SUBAPPLICATION Button_IXA_OR_AX_BG (* Button (IXA) ODER AX-Eingang, Ergebnis als Hintergrundfarbe (Gruen/Weiss) und AX-Ausgang *)
  (* Standard: 61499-2; Description: Copyright (c) 2026 Meisterschulen am Ostbahnhof This program and the accompanying materials are made available under the terms of the Eclipse Public License 2.0 which is available at https://www.eclipse.org/legal/epl-2.0/ SPDX-License-Identifier: EPL-2.0 *)
  (* Version 1.0, 2026-10-31, Franz Höpfinger, Meisterschulen am Ostbahnhof, Aus Getreidehacke func/Manual/ManFuncTast0 in MyLib::sys verschoben und umbenannt, INIT/INITO/QI/QO ergaenzt. *)
  PACKAGE MyLib::sys;
  IMPORT isobus::UT::Q::const::IDs::ID_NULL;
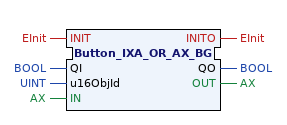
  EVENT_INPUT
    INIT : EInit; (* Initialization Request *)
  END_EVENT
  EVENT_OUTPUT
    INITO : EInit; (* Initialization Confirm *)
  END_EVENT
  VAR_INPUT
    QI : BOOL := TRUE; (* Quality Input - TRUE to enable service *)
    u16ObjId : UINT := ID_NULL; (* Object ID Button *)
  END_VAR
  VAR_OUTPUT
    QO : BOOL; (* Quality Output - TRUE if service executed successfully *)
  END_VAR
  SOCKETS
    IN : adapter::types::unidirectional::AX; (* zusaetzlicher Eingang, ODER mit Button *)
  END_SOCKETS
  PLUGS
    OUT : adapter::types::unidirectional::AX; (* Button ODER IN *)
  END_PLUGS
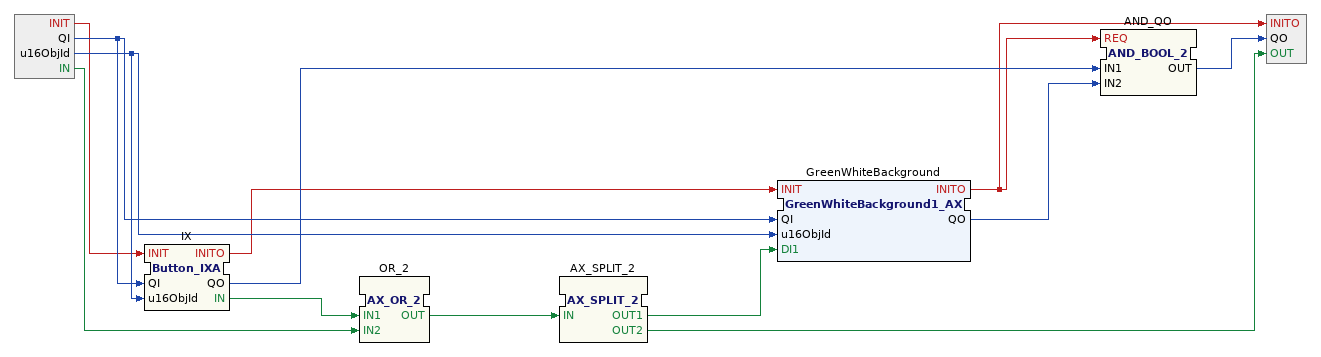
  FBS
    IX : isobus::UT::io::Button::Button_IXA;
    OR_2 : adapter::booleanOperators::AX_OR_2;
    AX_SPLIT_2 : adapter::events::unidirectional::AX_SPLIT_2;
    AND_QO : iec61131::booleanOperators::AND_BOOL_2;
  END_FBS
  SUBAPPS
    GreenWhiteBackground : MyLib::sys::GreenWhiteBackground1_AX;
  END_SUBAPPS
  EVENT_CONNECTIONS
    INIT TO IX.INIT;
    IX.INITO TO GreenWhiteBackground.INIT;
    GreenWhiteBackground.INITO TO INITO;
    GreenWhiteBackground.INITO TO AND_QO.REQ;
  END_CONNECTIONS
  DATA_CONNECTIONS
    QI TO IX.QI;
    QI TO GreenWhiteBackground.QI;
    u16ObjId TO IX.u16ObjId;
    u16ObjId TO GreenWhiteBackground.u16ObjId;
    IX.QO TO AND_QO.IN1;
    GreenWhiteBackground.QO TO AND_QO.IN2;
    AND_QO.OUT TO QO;
  END_CONNECTIONS
  ADAPTER_CONNECTIONS
    IX.IN TO OR_2.IN1;
    IN TO OR_2.IN2;
    OR_2.OUT TO AX_SPLIT_2.IN;
    AX_SPLIT_2.OUT1 TO GreenWhiteBackground.DI1;
    AX_SPLIT_2.OUT2 TO OUT;
  END_CONNECTIONS
END_SUBAPPLICATION
